//{attribute 'qualified_only'}
VAR_GLOBAL
	fbPump			: ARRAY[0..E_Pump_List.last] OF FB_Pump	;
	arr_st_Pump		: ARRAY[0..E_Pump_List.last] OF ST_Pump	;
	eClientPump		: E_Pump_List:= E_Pump_List.P1001;//eNotSelected;
	eClientStirrer	: E_Pump_List:= E_Pump_List.eNotSelected;//eNotSelected;
	
	fbDosingPP1002: FB_DosingPump; //Detergent
	fbDosingPP1003: FB_DosingPump; //DisInfection

END_VAR

(* stored: Version 1.1.0.1, ProductVersion 3.1.4024.13
   GVL g_Pump: Id {69c0cc40-2ece-41e7-8a9e-2b2b6efe872a} *)
